        pointRx pInter
        paraItem pParaItem
          [0]
            bool bSafePoint
            ifItem iIfItem
              [0]
                bool bANDOR[2]
                num nSigIndex[3]
                num nSigType[3]
                num nValue[3]
            mdesc mMdesc = {accel=0.64, vel=8, leave=0}
            num nActionIndex = 8
            num nDelay
            num nMoveType = 1
            num nPercentage
            num nSigValue = 1
        pointRx pPointRx[2] = {x=644.234527, y=1.0658073, z=249.473106, rx=-0.711473, ry=134.458377, rz=1.533345, shoulder=lefty, elbow=epositive, wrist=wpositive}
        string sID
      [27]
        bool bMarked
        jointRx jJointRx = {j1=-1.639045, j2=12.402747, j3=111.595585, j4=2.517874, j5=-30.594648, j6=-1.669011}
        pointRx pInter
        paraItem pParaItem
          [0]
            bool bSafePoint
            ifItem iIfItem
              [0]
                bool bANDOR[2]
                num nSigIndex[3]
                num nSigType[3]
                num nValue[3]
            mdesc mMdesc
            num nActionIndex = 10
            num nDelay = 5
            num nMoveType = 4
            num nPercentage
            num nSigValue
        pointRx pPointRx[2] = {x=594.549819, y=30.770866, z=171.45682, rx=-40.410864, ry=94.502866, rz=40.920287, shoulder=lefty, elbow=epositive, wrist=wnegative}
        string sID
      [28]
        bool bMarked
        jointRx jJointRx = {j1=-1.639045, j2=12.402747, j3=111.595585, j4=2.517874, j5=-30.594648, j6=-1.669011}
        pointRx pInter
        paraItem pParaItem
          [0]
            bool bSafePoint
            ifItem iIfItem
              [0]
                bool bANDOR[2]
                num nSigIndex[3]
                num nSigType[3]
                num nValue[3]
            mdesc mMdesc
            num nActionIndex = 10
            num nDelay = 0.5
            num nMoveType = 7
            num nPercentage
            num nSigValue
        pointRx pPointRx[2] = {x=594.549819, y=30.770866, z=171.45682, rx=-40.410864, ry=94.502866, rz=40.920287, shoulder=lefty, elbow=epositive, wrist=wnegative}
        string sID
      [29]
        bool bMarked
        jointRx jJointRx = {j1=-1.639045, j2=12.402747, j3=111.595585, j4=2.517874, j5=-30.594648, j6=-1.669011}
        pointRx pInter
        paraItem pParaItem
          [0]
            bool bSafePoint
            ifItem iIfItem
              [0]
                bool bANDOR[2]
                num nSigIndex[3]
                num nSigType[3]
                num nValue[3]
            mdesc mMdesc
            num nActionIndex = 9
            num nDelay = 5
            num nMoveType = 3
            num nPercentage
            num nSigValue = 1
        pointRx pPointRx[2] = {x=594.549819, y=30.770866, z=171.45682, rx=-40.410864, ry=94.502866, rz=40.920287, shoulder=lefty, elbow=epositive, wrist=wnegative}
        string sID
      [30]
        bool bMarked
        jointRx jJointRx = {j1=-3.707235, j2=5.145109, j3=114.936454, j4=-3.348646, j5=-32.0505381, j6=3.0814534}
        pointRx pInter
        paraItem pParaItem
          [0]
            bool bSafePoint
            ifItem iIfItem
              [0]
                bool bANDOR[2]
                num nSigIndex[3]
                num nSigType[3]
                num nValue[3]
            mdesc mMdesc = {leave=0}
            num nActionIndex = 9
            num nDelay = 5
            num nMoveType
            num nPercentage
            num nSigValue = 1
        pointRx pPointRx[2] = {x=558.0371815, y=17.0536556, z=213.621269, rx=45.0717683, ry=87.275085, rz=-44.921572, shoulder=lefty, elbow=epositive, wrist=wnegative}
        string sID
      [31]
        bool bMarked
        jointRx jJointRx = {j1=-6.48941, j2=24.903525, j3=114.355019, j4=-4.0836864, j5=-76.926301, j6=7.315242}
        pointRx pInter
        paraItem pParaItem
          [0]
            bool bSafePoint
            ifItem iIfItem
              [0]
                bool bANDOR[2]
                num nSigIndex[3]
                num nSigType[3]
                num nValue[3]
            mdesc mMdesc
            num nActionIndex = 1
            num nDelay = 5
            num nMoveType = 6
            num nPercentage
            num nSigValue = 1
        pointRx pPointRx[2] = {x=597.341422, y=-10.642707, z=109.749181, rx=3.827982, ry=62.369719, rz=-0.00899232, shoulder=lefty, elbow=epositive, wrist=wnegative}
        string sID
      [32]
        bool bMarked
        jointRx jJointRx = {j1=-6.48941, j2=24.903525, j3=114.355019, j4=-4.0836864, j5=-76.926301, j6=7.315242}
        pointRx pInter
        paraItem pParaItem
          [0]
            bool bSafePoint
            ifItem iIfItem
              [0]
                bool bANDOR[2]
                num nSigIndex[3]
                num nSigType[3]
                num nValue[3]
            mdesc mMdesc
            num nActionIndex = 1
            num nDelay = 5
            num nMoveType = 5
            num nPercentage
            num nSigValue = 1
        pointRx pPointRx[2] = {x=597.341422, y=-10.642707, z=109.749181, rx=3.827982, ry=62.369719, rz=-0.00899232, shoulder=lefty, elbow=epositive, wrist=wnegative}
        string sID
      [33]
        bool bMarked
        jointRx jJointRx = {j1=-6.48941, j2=24.903525, j3=114.355019, j4=-4.0836864, j5=-76.926301, j6=7.315242}
        pointRx pInter
        paraItem pParaItem
          [0]
            bool bSafePoint
            ifItem iIfItem
              [0]
                bool bANDOR[2]
                num nSigIndex[3]
                num nSigType[3]
                num nValue[3]
            mdesc mMdesc
            num nActionIndex = 10
            num nDelay = 5
            num nMoveType = 4
            num nPercentage
            num nSigValue = 1
        pointRx pPointRx[2] = {x=597.341422, y=-10.642707, z=109.749181, rx=3.827982, ry=62.369719, rz=-0.00899232, shoulder=lefty, elbow=epositive, wrist=wnegative}
        string sID
      [34]
        bool bMarked
        jointRx jJointRx = {j1=-6.48941, j2=24.903525, j3=114.355019, j4=-4.0836864, j5=-76.926301, j6=7.315242}
        pointRx pInter
        paraItem pParaItem
          [0]
            bool bSafePoint
            ifItem iIfItem
              [0]
                bool bANDOR[2]
                num nSigIndex[3]
                num nSigType[3]
                num nValue[3]
            mdesc mMdesc
            num nActionIndex = 8
            num nDelay = 5
            num nMoveType = 3
            num nPercentage
            num nSigValue = 1
        pointRx pPointRx[2] = {x=597.341422, y=-10.642707, z=109.749181, rx=3.827982, ry=62.369719, rz=-0.00899232, shoulder=lefty, elbow=epositive, wrist=wnegative}
        string sID
      [35]
        bool bMarked
        jointRx jJointRx = {j1=-3.703679, j2=18.38504, j3=121.854236, j4=-2.248579, j5=-52.181366, j6=1.621257}
        pointRx pInter
        paraItem pParaItem
          [0]
            bool bSafePoint
            ifItem iIfItem
              [0]
                bool bANDOR[2]
                num nSigIndex[3]
                num nSigType[3]
                num nValue[3]
            mdesc mMdesc = {accel=0.64, vel=8, leave=0}
            num nActionIndex = 8
            num nDelay = 5
            num nMoveType = 1
            num nPercentage
            num nSigValue = 1
        pointRx pPointRx[2] = {x=558.0333709, y=17.0881425, z=79.950444, rx=45.0849978, ry=87.280462, rz=-44.934765, shoulder=lefty, elbow=epositive, wrist=wnegative}
        string sID
      [36]
        bool bMarked
        jointRx jJointRx = {j1=-6.48941, j2=24.903525, j3=114.355019, j4=-4.0836864, j5=-76.926301, j6=7.315242}
        pointRx pInter
        paraItem pParaItem
          [0]
            bool bSafePoint
            ifItem iIfItem
              [0]
                bool bANDOR[2]
                num nSigIndex[3]
                num nSigType[3]
                num nValue[3]
            mdesc mMdesc
            num nActionIndex = 10
            num nDelay = 1
            num nMoveType = 4
            num nPercentage
            num nSigValue
        pointRx pPointRx[2] = {x=597.341422, y=-10.642707, z=109.749181, rx=3.827982, ry=62.369719, rz=-0.00899232, shoulder=lefty, elbow=epositive, wrist=wnegative}
        string sID
      [37]
        bool bMarked
        jointRx jJointRx = {j1=-6.48941, j2=24.903525, j3=114.355019, j4=-4.0836864, j5=-76.926301, j6=7.315242}
        pointRx pInter
        paraItem pParaItem
          [0]
            bool bSafePoint
            ifItem iIfItem
              [0]
                bool bANDOR[2]
                num nSigIndex[3]
                num nSigType[3]
                num nValue[3]
            mdesc mMdesc
            num nActionIndex = 9
            num nDelay = 1
            num nMoveType = 3
            num nPercentage
            num nSigValue = 1
        pointRx pPointRx[2] = {x=597.341422, y=-10.642707, z=109.749181, rx=3.827982, ry=62.369719, rz=-0.00899232, shoulder=lefty, elbow=epositive, wrist=wnegative}
        string sID
      [38]
        bool bMarked
        jointRx jJointRx = {j1=-1.639045, j2=12.402747, j3=111.595585, j4=2.517874, j5=-30.594648, j6=-1.669011}
        pointRx pInter
        paraItem pParaItem
          [0]
            bool bSafePoint
            ifItem iIfItem
              [0]
                bool bANDOR[2]
                num nSigIndex[3]
                num nSigType[3]
                num nValue[3]
            mdesc mMdesc
            num nActionIndex = 1
            num nDelay = 5
            num nMoveType = 6
            num nPercentage
            num nSigValue
        pointRx pPointRx[2] = {x=594.549819, y=30.770866, z=171.45682, rx=-40.410864, ry=94.502866, rz=40.920287, shoulder=lefty, elbow=epositive, wrist=wnegative}
        string sID
      [39]
        bool bMarked
        jointRx jJointRx = {j1=-1.639045, j2=12.402747, j3=111.595585, j4=2.517874, j5=-30.594648, j6=-1.669011}
        pointRx pInter
        paraItem pParaItem
          [0]
            bool bSafePoint
            ifItem iIfItem
              [0]
                bool bANDOR[2]
                num nSigIndex[3]
                num nSigType[3]
                num nValue[3]
            mdesc mMdesc
            num nActionIndex = 1
            num nDelay = 5
            num nMoveType = 5
            num nPercentage
            num nSigValue
        pointRx pPointRx[2] = {x=594.549819, y=30.770866, z=171.45682, rx=-40.410864, ry=94.502866, rz=40.920287, shoulder=lefty, elbow=epositive, wrist=wnegative}
        string sID
      [40]
        bool bMarked
        jointRx jJointRx = {j1=-6.652009, j2=-3.724795, j3=129.0452396, j4=-6.346388, j5=-34.648815, j6=4.794651}
        pointRx pInter
        paraItem pParaItem
          [0]
            bool bSafePoint
            ifItem iIfItem
              [0]
                bool bANDOR[2]
                num nSigIndex[3]
                num nSigType[3]
                num nValue[3]
            mdesc mMdesc
            num nActionIndex = 1
            num nDelay = 5
            num nMoveType
            num nPercentage
            num nSigValue
        pointRx pPointRx[2] = {x=472.315715, y=1.582801, z=176.932517, rx=-74.682061, ry=93.16048, rz=74.323701, shoulder=lefty, elbow=epositive, wrist=wnegative}
        string sID
      [41]
        bool bMarked
        jointRx jJointRx = {j1=-1.639045, j2=12.402747, j3=111.595585, j4=2.517874, j5=-30.594648, j6=-1.669011}
        pointRx pInter
        paraItem pParaItem
          [0]
            bool bSafePoint
            ifItem iIfItem
              [0]
                bool bANDOR[2]
                num nSigIndex[3]
                num nSigType[3]
                num nValue[3]
            mdesc mMdesc
            num nActionIndex = 11
            num nDelay = 5
            num nMoveType = 4
            num nPercentage
            num nSigValue = 1
        pointRx pPointRx[2] = {x=594.549819, y=30.770866, z=171.45682, rx=-40.410864, ry=94.502866, rz=40.920287, shoulder=lefty, elbow=epositive, wrist=wnegative}
        string sID
      [42]
        bool bMarked
        jointRx jJointRx = {j1=-1.639045, j2=12.402747, j3=111.595585, j4=2.517874, j5=-30.594648, j6=-1.669011}
        pointRx pInter
        paraItem pParaItem
          [0]
            bool bSafePoint
            ifItem iIfItem
              [0]
                bool bANDOR[2]
                num nSigIndex[3]
                num nSigType[3]
                num nValue[3]
            mdesc mMdesc
            num nActionIndex = 10
            num nDelay = 5
            num nMoveType = 3
            num nPercentage
            num nSigValue
        pointRx pPointRx[2] = {x=594.549819, y=30.770866, z=171.45682, rx=-40.410864, ry=94.502866, rz=40.920287, shoulder=lefty, elbow=epositive, wrist=wnegative}
        string sID
      [43]
        bool bMarked
        jointRx jJointRx = {j1=-1.639045, j2=12.402747, j3=111.595585, j4=2.517874, j5=-30.594648, j6=-1.669011}
        pointRx pInter
        paraItem pParaItem
          [0]
            bool bSafePoint
            ifItem iIfItem
              [0]
                bool bANDOR[2]
                num nSigIndex[3]
                num nSigType[3]
                num nValue[3]
            mdesc mMdesc
            num nActionIndex = 9
            num nDelay = 5
            num nMoveType = 4
            num nPercentage
            num nSigValue
        pointRx pPointRx[2] = {x=594.549819, y=30.770866, z=171.45682, rx=-40.410864, ry=94.502866, rz=40.920287, shoulder=lefty, elbow=epositive, wrist=wnegative}
        string sID
      [44]
        bool bMarked
        jointRx jJointRx = {j1=-1.639045, j2=12.402747, j3=111.595585, j4=2.517874, j5=-30.594648, j6=-1.669011}
        pointRx pInter
        paraItem pParaItem
          [0]
            bool bSafePoint
            ifItem iIfItem
              [0]
                bool bANDOR[2]
                num nSigIndex[3]
                num nSigType[3]
                num nValue[3]
            mdesc mMdesc
            num nActionIndex = 11
            num nDelay = 5
            num nMoveType = 4
            num nPercentage
            num nSigValue
        pointRx pPointRx[2] = {x=594.549819, y=30.770866, z=171.45682, rx=-40.410864, ry=94.502866, rz=40.920287, shoulder=lefty, elbow=epositive, wrist=wnegative}
        string sID
    string sID
  [04 sls]
    num nFrameIndex
    num nMoveID
    num nToolIndex
    pointItem pPointItem[96]
      [0]
        bool bMarked
        jointRx jJointRx = {j1=-2.594987, j2=-12.391258, j3=136.392534, j4=0.644488, j5=-30.575639, j6=-0.113504}
        pointRx pInter
        paraItem pParaItem
          [0]
            bool bSafePoint
            ifItem iIfItem
              [0]
                bool bANDOR[2]
                num nSigIndex[3]
                num nSigType[3]
                num nValue[3]
            mdesc mMdesc
            num nActionIndex = 11
            num nDelay
            num nMoveType = 4
            num nPercentage
            num nSigValue
        pointRx pPointRx[2] = {x=412.772469, y=30.77087, z=171.456836, rx=-40.418431, ry=94.503508, rz=40.927655, shoulder=lefty, elbow=epositive, wrist=wnegative}
        string sID
      [1]
        bool bMarked
        jointRx jJointRx = {j1=-2.594987, j2=-12.391258, j3=136.392534, j4=0.644488, j5=-30.575639, j6=-0.113504}
        pointRx pInter
        paraItem pParaItem
          [0]
            bool bSafePoint
            ifItem iIfItem
              [0]
                bool bANDOR[2]
                num nSigIndex[3]
                num nSigType[3]
                num nValue[3]
            mdesc mMdesc
            num nActionIndex = 9
            num nDelay
            num nMoveType = 4
            num nPercentage
            num nSigValue = 1
        pointRx pPointRx[2] = {x=412.772469, y=30.77087, z=171.456836, rx=-40.418431, ry=94.503508, rz=40.927655, shoulder=lefty, elbow=epositive, wrist=wnegative}
        string sID
      [2]
        bool bMarked
        jointRx jJointRx = {j1=-6.648888, j2=-3.725245, j3=129.0447888, j4=-6.34617, j5=-34.648619, j6=4.79455}
        pointRx pInter
        paraItem pParaItem
          [0]
            bool bSafePoint
            ifItem iIfItem
              [0]
                bool bANDOR[2]
                num nSigIndex[3]
                num nSigType[3]
                num nValue[3]
            mdesc mMdesc
            num nActionIndex
            num nDelay
            num nMoveType
            num nPercentage
            num nSigValue
        pointRx pPointRx[2] = {x=472.316162, y=1.608216, z=176.938999, rx=-74.680314, ry=93.157419, rz=74.321932, shoulder=lefty, elbow=epositive, wrist=wnegative}
        string sID
      [3]
        bool bMarked
        jointRx jJointRx = {j1=-6.652767, j2=20.832827, j3=135.880999, j4=-3.946436, j5=-65.929599, j6=1.179192}
        pointRx pInter
        paraItem pParaItem
          [0]
            bool bSafePoint
            ifItem iIfItem
              [0]
                bool bANDOR[2]
                num nSigIndex[3]
                num nSigType[3]
                num nValue[3]
            mdesc mMdesc
            num nActionIndex
            num nDelay
            num nMoveType
            num nPercentage
            num nSigValue
        pointRx pPointRx[2] = {x=472.315383, y=1.575881, z=5.379837, rx=-74.70962, ry=93.161274, rz=74.351748, shoulder=lefty, elbow=epositive, wrist=wnegative}
        string sID
      [4]
        bool bMarked
        jointRx jJointRx = {j1=-3.751907, j2=40.467467, j3=104.535855, j4=-3.0941224, j5=-89.629669, j6=3.053905}
        pointRx pInter
        paraItem pParaItem
          [0]
            bool bSafePoint
            ifItem iIfItem
              [0]
                bool bANDOR[2]
                num nSigIndex[3]
                num nSigType[3]
                num nValue[3]
            mdesc mMdesc
            num nActionIndex
            num nDelay
            num nMoveType
            num nPercentage
            num nSigValue
        pointRx pPointRx[2] = {x=653.977922, y=12.630674, z=31.914071, rx=-0.00926733, ry=55.431846, rz=0.910662, shoulder=lefty, elbow=epositive, wrist=wnegative}
        string sID
      [5]
        bool bMarked
        jointRx jJointRx = {j1=-1.639045, j2=12.402747, j3=111.595585, j4=2.517874, j5=-30.594648, j6=-1.669011}
        pointRx pInter
        paraItem pParaItem
          [0]
            bool bSafePoint
            ifItem iIfItem
              [0]
                bool bANDOR[2]
                num nSigIndex[3]
                num nSigType[3]
                num nValue[3]
            mdesc mMdesc
            num nActionIndex = 1
            num nDelay
            num nMoveType = 6
            num nPercentage
            num nSigValue = 1
        pointRx pPointRx[2] = {x=594.549819, y=30.770866, z=171.45682, rx=-40.410864, ry=94.502866, rz=40.920287, shoulder=lefty, elbow=epositive, wrist=wnegative}
        string sID
      [6]
        bool bMarked
        jointRx jJointRx = {j1=-1.639045, j2=12.402747, j3=111.595585, j4=2.517874, j5=-30.594648, j6=-1.669011}
        pointRx pInter
        paraItem pParaItem
          [0]
            bool bSafePoint
            ifItem iIfItem
              [0]
                bool bANDOR[2]
                num nSigIndex[3]
                num nSigType[3]
                num nValue[3]
            mdesc mMdesc
            num nActionIndex = 1
            num nDelay
            num nMoveType = 5
            num nPercentage
            num nSigValue = 1
        pointRx pPointRx[2] = {x=594.549819, y=30.770866, z=171.45682, rx=-40.410864, ry=94.502866, rz=40.920287, shoulder=lefty, elbow=epositive, wrist=wnegative}
        string sID
      [7]
        bool bMarked
        jointRx jJointRx = {j1=-1.639045, j2=12.402747, j3=111.595585, j4=2.517874, j5=-30.594648, j6=-1.669011}
        pointRx pInter
        paraItem pParaItem
          [0]
            bool bSafePoint
            ifItem iIfItem
              [0]
                bool bANDOR[2]
                num nSigIndex[3]
                num nSigType[3]
                num nValue[3]
            mdesc mMdesc
            num nActionIndex = 10
            num nDelay
            num nMoveType = 4
            num nPercentage
            num nSigValue = 1
        pointRx pPointRx[2] = {x=594.549819, y=30.770866, z=171.45682, rx=-40.410864, ry=94.502866, rz=40.920287, shoulder=lefty, elbow=epositive, wrist=wnegative}
        string sID
      [8]
        bool bMarked
        jointRx jJointRx = {j1=-1.639045, j2=12.402747, j3=111.595585, j4=2.517874, j5=-30.594648, j6=-1.669011}
        pointRx pInter
        paraItem pParaItem
          [0]
            bool bSafePoint
            ifItem iIfItem
              [0]
                bool bANDOR[2]
                num nSigIndex[3]
                num nSigType[3]
                num nValue[3]
            mdesc mMdesc
            num nActionIndex = 8
            num nDelay
            num nMoveType = 3
            num nPercentage
            num nSigValue = 1
        pointRx pPointRx[2] = {x=594.549819, y=30.770866, z=171.45682, rx=-40.410864, ry=94.502866, rz=40.920287, shoulder=lefty, elbow=epositive, wrist=wnegative}
        string sID
      [9]
        bool bMarked
        jointRx jJointRx = {j1=-1.639045, j2=12.402747, j3=111.595585, j4=2.517874, j5=-30.594648, j6=-1.669011}
        pointRx pInter
        paraItem pParaItem
          [0]
            bool bSafePoint
            ifItem iIfItem
              [0]
                bool bANDOR[2]
                num nSigIndex[3]
                num nSigType[3]
                num nValue[3]
            mdesc mMdesc
            num nActionIndex = 8
            num nDelay = 2
            num nMoveType = 7
            num nPercentage
            num nSigValue = 1
        pointRx pPointRx[2] = {x=594.549819, y=30.770866, z=171.45682, rx=-40.410864, ry=94.502866, rz=40.920287, shoulder=lefty, elbow=epositive, wrist=wnegative}
        string sID
      [10]
        bool bMarked
        jointRx jJointRx = {j1=-1.639045, j2=12.402747, j3=111.595585, j4=2.517874, j5=-30.594648, j6=-1.669011}
        pointRx pInter
        paraItem pParaItem
          [0]
            bool bSafePoint
            ifItem iIfItem
              [0]
                bool bANDOR[2]
                num nSigIndex[3]
                num nSigType[3]
                num nValue[3]
            mdesc mMdesc
            num nActionIndex = 10
            num nDelay = 5
            num nMoveType = 4
            num nPercentage
            num nSigValue
        pointRx pPointRx[2] = {x=594.549819, y=30.770866, z=171.45682, rx=-40.410864, ry=94.502866, rz=40.920287, shoulder=lefty, elbow=epositive, wrist=wnegative}
        string sID
      [11]
        bool bMarked
        jointRx jJointRx = {j1=-1.639045, j2=12.402747, j3=111.595585, j4=2.517874, j5=-30.594648, j6=-1.669011}
        pointRx pInter
        paraItem pParaItem
          [0]
            bool bSafePoint
            ifItem iIfItem
              [0]
                bool bANDOR[2]
                num nSigIndex[3]
                num nSigType[3]
                num nValue[3]
            mdesc mMdesc
            num nActionIndex = 10
            num nDelay = 0.5
            num nMoveType = 7
            num nPercentage
            num nSigValue
        pointRx pPointRx[2] = {x=594.549819, y=30.770866, z=171.45682, rx=-40.410864, ry=94.502866, rz=40.920287, shoulder=lefty, elbow=epositive, wrist=wnegative}
        string sID
      [12]
        bool bMarked
        jointRx jJointRx = {j1=-1.639045, j2=12.402747, j3=111.595585, j4=2.517874, j5=-30.594648, j6=-1.669011}
        pointRx pInter
        paraItem pParaItem
          [0]
            bool bSafePoint
            ifItem iIfItem
              [0]
                bool bANDOR[2]
                num nSigIndex[3]
                num nSigType[3]
                num nValue[3]
            mdesc mMdesc
            num nActionIndex = 9
            num nDelay = 5
            num nMoveType = 3
            num nPercentage
            num nSigValue = 1
        pointRx pPointRx[2] = {x=594.549819, y=30.770866, z=171.45682, rx=-40.410864, ry=94.502866, rz=40.920287, shoulder=lefty, elbow=epositive, wrist=wnegative}
        string sID
      [13]
        bool bMarked
        jointRx jJointRx = {j1=-6.995994, j2=22.295183, j3=133.491067, j4=-6.412947, j5=-89.696299, j6=3.773786}
        pointRx pInter
        paraItem pParaItem
          [0]
            bool bSafePoint
            ifItem iIfItem
              [0]
                bool bANDOR[2]
                num nSigIndex[3]
                num nSigType[3]
                num nValue[3]
            mdesc mMdesc
            num nActionIndex
            num nDelay
            num nMoveType
            num nPercentage
            num nSigValue
        pointRx pPointRx[2] = {x=480.297234, y=2.689037, z=45.892011, rx=-0.0295899, ry=66.250693, rz=0.93735, shoulder=lefty, elbow=epositive, wrist=wnegative}
        string sID
      [14]
        bool bMarked
        jointRx jJointRx = {j1=-3.631024, j2=-1.590232, j3=111.256847, j4=-19.293027, j5=-7.965925, j6=19.0488477}
        pointRx pInter
        paraItem pParaItem
          [0]
            bool bSafePoint
            ifItem iIfItem
              [0]
                bool bANDOR[2]
                num nSigIndex[3]
                num nSigType[3]
                num nValue[3]
            mdesc mMdesc = {leave=1}
            num nActionIndex
            num nDelay
            num nMoveType = 1
            num nPercentage
            num nSigValue
        pointRx pPointRx[2] = {x=538.454635, y=20.519182, z=260.791216, rx=-4.395762, ry=102.166176, rz=4.98921, shoulder=lefty, elbow=epositive, wrist=wnegative}
        string sID
      [15]
        bool bMarked
        jointRx jJointRx = {j1=-2.334364, j2=-5.268397, j3=112.836865, j4=-1.917467, j5=-5.341213, j6=2.362596}
        pointRx pInter
        paraItem pParaItem
          [0]
            bool bSafePoint
            ifItem iIfItem
              [0]
                bool bANDOR[2]
                num nSigIndex[3]
                num nSigType[3]
                num nValue[3]
            mdesc mMdesc = {leave=1}
            num nActionIndex = 1
            num nDelay
            num nMoveType = 6
            num nPercentage
            num nSigValue = 1
        pointRx pPointRx[2] = {x=515.505365, y=29.338734, z=273.736407, rx=-9.827138, ry=102.415174, rz=10.549826, shoulder=lefty, elbow=epositive, wrist=wnegative}
        string sID
      [16]
        bool bMarked
        jointRx jJointRx = {j1=-2.334364, j2=-5.268397, j3=112.836865, j4=-1.917467, j5=-5.341213, j6=2.362596}
        pointRx pInter
        paraItem pParaItem
          [0]
            bool bSafePoint
            ifItem iIfItem
              [0]
                bool bANDOR[2]
                num nSigIndex[3]
                num nSigType[3]
                num nValue[3]
            mdesc mMdesc = {leave=1}
            num nActionIndex = 1
            num nDelay
            num nMoveType = 5
            num nPercentage
            num nSigValue = 1
        pointRx pPointRx[2] = {x=515.505365, y=29.338734, z=273.736407, rx=-9.827138, ry=102.415174, rz=10.549826, shoulder=lefty, elbow=epositive, wrist=wnegative}
        string sID
      [17]
        bool bMarked
        jointRx jJointRx = {j1=-1.639045, j2=12.402747, j3=111.595585, j4=2.517874, j5=-30.594648, j6=-1.669011}
        pointRx pInter
        paraItem pParaItem
          [0]
            bool bSafePoint
            ifItem iIfItem
              [0]
                bool bANDOR[2]
                num nSigIndex[3]
                num nSigType[3]
                num nValue[3]
            mdesc mMdesc
            num nActionIndex = 10
            num nDelay
            num nMoveType = 4
            num nPercentage
            num nSigValue = 1
        pointRx pPointRx[2] = {x=594.549819, y=30.770866, z=171.45682, rx=-40.410864, ry=94.502866, rz=40.920287, shoulder=lefty, elbow=epositive, wrist=wnegative}
        string sID
      [18]
        bool bMarked
        jointRx jJointRx = {j1=-1.639045, j2=12.402747, j3=111.595585, j4=2.517874, j5=-30.594648, j6=-1.669011}
        pointRx pInter
        paraItem pParaItem
          [0]
            bool bSafePoint
            ifItem iIfItem
              [0]
                bool bANDOR[2]
                num nSigIndex[3]
                num nSigType[3]
                num nValue[3]
            mdesc mMdesc
            num nActionIndex = 8
            num nDelay
            num nMoveType = 3
            num nPercentage
            num nSigValue = 1
        pointRx pPointRx[2] = {x=594.549819, y=30.770866, z=171.45682, rx=-40.410864, ry=94.502866, rz=40.920287, shoulder=lefty, elbow=epositive, wrist=wnegative}
        string sID
      [19]
        bool bMarked
        jointRx jJointRx = {j1=-1.639045, j2=12.402747, j3=111.595585, j4=2.517874, j5=-30.594648, j6=-1.669011}
        pointRx pInter
        paraItem pParaItem
          [0]
            bool bSafePoint
            ifItem iIfItem
              [0]
                bool bANDOR[2]
                num nSigIndex[3]
                num nSigType[3]
                num nValue[3]
            mdesc mMdesc
            num nActionIndex = 8
            num nDelay = 0.8
            num nMoveType = 7
            num nPercentage
            num nSigValue = 1
        pointRx pPointRx[2] = {x=594.549819, y=30.770866, z=171.45682, rx=-40.410864, ry=94.502866, rz=40.920287, shoulder=lefty, elbow=epositive, wrist=wnegative}
        string sID
      [20]
        bool bMarked
        jointRx jJointRx = {j1=-1.639045, j2=12.402747, j3=111.595585, j4=2.517874, j5=-30.594648, j6=-1.669011}
        pointRx pInter
        paraItem pParaItem
          [0]
            bool bSafePoint
            ifItem iIfItem
              [0]
                bool bANDOR[2]
                num nSigIndex[3]
                num nSigType[3]
                num nValue[3]
            mdesc mMdesc
            num nActionIndex = 10
            num nDelay = 5
            num nMoveType = 4
            num nPercentage
            num nSigValue
        pointRx pPointRx[2] = {x=594.549819, y=30.770866, z=171.45682, rx=-40.410864, ry=94.502866, rz=40.920287, shoulder=lefty, elbow=epositive, wrist=wnegative}
        string sID
      [21]
        bool bMarked
        jointRx jJointRx = {j1=-1.639045, j2=12.402747, j3=111.595585, j4=2.517874, j5=-30.594648, j6=-1.669011}
        pointRx pInter
        paraItem pParaItem
          [0]
            bool bSafePoint
            ifItem iIfItem
              [0]
                bool bANDOR[2]
                num nSigIndex[3]
                num nSigType[3]
                num nValue[3]
            mdesc mMdesc
            num nActionIndex = 10
            num nDelay = 0.5
            num nMoveType = 7
            num nPercentage
            num nSigValue
        pointRx pPointRx[2] = {x=594.549819, y=30.770866, z=171.45682, rx=-40.410864, ry=94.502866, rz=40.920287, shoulder=lefty, elbow=epositive, wrist=wnegative}
        string sID
      [22]
        bool bMarked
        jointRx jJointRx = {j1=-1.639045, j2=12.402747, j3=111.595585, j4=2.517874, j5=-30.594648, j6=-1.669011}
        pointRx pInter
        paraItem pParaItem
          [0]
            bool bSafePoint
            ifItem iIfItem
              [0]
                bool bANDOR[2]
                num nSigIndex[3]
                num nSigType[3]
                num nValue[3]
            mdesc mMdesc
            num nActionIndex = 9
            num nDelay = 5
            num nMoveType = 3
            num nPercentage
            num nSigValue = 1
        pointRx pPointRx[2] = {x=594.549819, y=30.770866, z=171.45682, rx=-40.410864, ry=94.502866, rz=40.920287, shoulder=lefty, elbow=epositive, wrist=wnegative}
        string sID
      [23]
        bool bMarked
        jointRx jJointRx = {j1=-3.587733, j2=23.639281, j3=117.919343, j4=-3.340268, j5=-74.590591, j6=2.335421}
        pointRx pInter
        paraItem pParaItem
          [0]
            bool bSafePoint
            ifItem iIfItem
              [0]
                bool bANDOR[2]
                num nSigIndex[3]
                num nSigType[3]
                num nValue[3]
            mdesc mMdesc
            num nActionIndex = 9
            num nDelay = 5
            num nMoveType
            num nPercentage
            num nSigValue = 1
        pointRx pPointRx[2] = {x=578.894359, y=19.429807, z=95.481067, rx=0.212509, ry=67.0312458, rz=-0.1502, shoulder=lefty, elbow=epositive, wrist=wnegative}
        string sID
      [24]
        bool bMarked
        jointRx jJointRx = {j1=-2.687248, j2=16.117165, j3=122.304638, j4=-0.487867, j5=-66.528565, j6=1.978834}
        pointRx pInter
        paraItem pParaItem
          [0]
            bool bSafePoint
            ifItem iIfItem
              [0]
                bool bANDOR[2]
                num nSigIndex[3]
                num nSigType[3]
                num nValue[3]
            mdesc mMdesc
            num nActionIndex = 1
            num nDelay = 5
            num nMoveType = 6
            num nPercentage
            num nSigValue = 1
        pointRx pPointRx[2] = {x=546.855577, y=25.169852, z=121.450925, rx=6.745985, ry=71.76392, rz=-5.460967, shoulder=lefty, elbow=epositive, wrist=wnegative}
        string sID
      [25]
        bool bMarked
        jointRx jJointRx = {j1=-2.687248, j2=16.117165, j3=122.304638, j4=-0.487867, j5=-66.528565, j6=1.978834}
        pointRx pInter
        paraItem pParaItem
          [0]
            bool bSafePoint
            ifItem iIfItem
              [0]
                bool bANDOR[2]
                num nSigIndex[3]
                num nSigType[3]
                num nValue[3]
            mdesc mMdesc
            num nActionIndex = 1
            num nDelay = 5
            num nMoveType = 5
            num nPercentage
            num nSigValue = 1
        pointRx pPointRx[2] = {x=546.855577, y=25.169852, z=121.450925, rx=6.745985, ry=71.76392, rz=-5.460967, shoulder=lefty, elbow=epositive, wrist=wnegative}
        string sID
      [26]
        bool bMarked
        jointRx jJointRx = {j1=-1.639045, j2=12.402747, j3=111.595585, j4=2.517874, j5=-30.594648, j6=-1.669011}
        pointRx pInter
        paraItem pParaItem
          [0]
            bool bSafePoint
            ifItem iIfItem
              [0]
                bool bANDOR[2]
                num nSigIndex[3]
                num nSigType[3]
                num nValue[3]
            mdesc mMdesc
            num nActionIndex = 10
            num nDelay
            num nMoveType = 4
            num nPercentage
            num nSigValue = 1
        pointRx pPointRx[2] = {x=594.549819, y=30.770866, z=171.45682, rx=-40.410864, ry=94.502866, rz=40.920287, shoulder=lefty, elbow=epositive, wrist=wnegative}
        string sID
      [27]
        bool bMarked
        jointRx jJointRx = {j1=-1.639045, j2=12.402747, j3=111.595585, j4=2.517874, j5=-30.594648, j6=-1.669011}
        pointRx pInter
        paraItem pParaItem
          [0]
            bool bSafePoint
            ifItem iIfItem
              [0]
                bool bANDOR[2]
                num nSigIndex[3]
                num nSigType[3]
                num nValue[3]
            mdesc mMdesc
            num nActionIndex = 8
            num nDelay
            num nMoveType = 3
            num nPercentage
            num nSigValue = 1
